TYPE ST_ITECH_SystemStatus :
STRUCT
	ON_OFF				: UDINT;
	SenseVolt			: REAL;
	Heartbeat			: UDINT;
	Timer_ON_OFF		: UDINT;
	RemoteSenseStatus	: UDINT;
	RemoteSenseLevel	: REAL;
	OutputRZero			: UDINT;
	MeasureCycle		: UDINT;
END_STRUCT
END_TYPE

(* stored: Version 1.1.0.1
   DUT ST_ITECH_SystemStatus: Id {7ac071da-9578-4fcd-9e35-fef6269e2dfb} *)
